Fanuc KAREL source: KA00226.KL

PROGRAM KA00226
%NOLOCKGROUP
VAR
  SRC: FILE
  DST: FILE
BEGIN
  DST = SRC
END KA00226
